// TIA Portal project "PLC_5_LINE5" (V18)

(* hardware
DEVICE "S7-1500/ET200MP station_1"  S7-1500 station
   slot 0: "Rail_0"  Rack  6ES7 590-1***0-0AA0
   slot 1: "PLC_1"  CPU 1511-1 PN  6ES7 511-1AK02-0AB0  V2.9
      slot 3: "CPU display_1"  6ES7591-1AA00-0AA0
      slot 32768: "PROFINET interface_1"  X1
         slot 32769: "Port_1"  X1 P1
         slot 32770: "Port_2"  X1 P2
      slot 34817: "Virtual CP interface port_1"  Virtual CP interface port  Virtual CP interface port
   slot 2: "DI 32x24VDC HF_1"  DI 32x24VDC HF  6ES7 521-1BL00-0AB0  V2.2
   slot 3: "DQ 32x24VDC/0.5A HF_1"  DQ 32x24VDC/0.5A HF  6ES7 522-1BL01-0AB0  V1.1
*)

// ===== PLC "PLC_1"  CPU 1511-1 PN =====

VAR_GLOBAL   // PLC tag table "Default tag table"
   "Tag_1" AT %I4.3 : Bool;
   "Tag_2" AT %I4.4 : Bool;
   "Tag_3" AT %I4.5 : Bool;
   "Tag_4" AT %I4.0 : Bool;
   "Tag_5" AT %I4.1 : Bool;
   "Tag_6" AT %I5.0 : Bool;
   "Tag_7" AT %I5.2 : Bool;
   "Tag_8" AT %I6.3 : Bool;
   "Tag_9" AT %I5.3 : Bool;
   "Tag_10" AT %I5.4 : Bool;
   "Tag_11" AT %I5.5 : Bool;
   "Tag_12" AT %I5.6 : Bool;
   "Tag_13" AT %I5.7 : Bool;
   "Tag_14" AT %I6.0 : Bool;
   "Tag_15" AT %I6.1 : Bool;
   "Tag_16" AT %I6.2 : Bool;
   "Tag_17" AT %Q1.6 : Bool;
   "Tag_18" AT %Q1.7 : Bool;
   "Tag_19" AT %Q2.0 : Bool;
   "Tag_20" AT %Q2.1 : Bool;
   "Tag_21" AT %Q2.2 : Bool;
   "Tag_22" AT %Q2.3 : Bool;
   "Tag_23" AT %I0.3 : Bool;
   "Tag_24" AT %I0.4 : Bool;
   "Tag_25" AT %I0.5 : Bool;
   "Tag_26" AT %I0.0 : Bool;
   "Tag_27" AT %I0.1 : Bool;
   "Tag_28" AT %I1.0 : Bool;
   "Tag_29" AT %I2.7 : Bool;
   "Tag_30" AT %I3.1 : Bool;
   "Tag_31" AT %I1.6 : Bool;
   "Tag_32" AT %I1.7 : Bool;
   "Tag_33" AT %I2.0 : Bool;
   "Tag_34" AT %I2.1 : Bool;
   "Tag_35" AT %I2.2 : Bool;
   "Tag_36" AT %I2.3 : Bool;
   "Tag_37" AT %I2.4 : Bool;
   "Tag_38" AT %I2.5 : Bool;
   "Tag_39" AT %I2.6 : Bool;
   "Tag_40" AT %I3.0 : Bool;
   "Tag_41" AT %Q0.4 : Bool;
   "Tag_42" AT %Q0.5 : Bool;
   "Tag_43" AT %Q0.6 : Bool;
   "Tag_44" AT %Q0.7 : Bool;
   "Tag_45" AT %Q1.0 : Bool;
   "Tag_46" AT %Q1.1 : Bool;
END_VAR

TYPE "typeTask"
   STRUCT
      station : Int;
      dwell_s : Int;
      crane : String[4];
      tank_name : String[10];
      prev : Int;
      next : Int;
      status : Int;
   END_STRUCT;
END_TYPE

TYPE "typeCraneData"
   STRUCT
      task_count : Int;
      tasks : Array[1..20] of "typeTask";
      cmd_send : Bool;
      sts_busy : Bool;
      sts_done : Bool;
      sts_step : Int;
      sts_state : Int;
      ls_at : Array[0..20] of Bool;
      ls_dip : Bool;
      ls_up : Bool;
      ls_mid : Bool;
      btn_start : Bool;
      mv_fwd : Bool;
      mv_rev : Bool;
      mv_up : Bool;
      mv_down : Bool;
      estop : Bool;
      auto : Bool;
      cmd_reset : Bool;
      cmd_stop : Bool;
      pos : Array[0..20] of Int;
   END_STRUCT;
END_TYPE

DATA_BLOCK "Crane8Data"   // DB1
{ S7_Optimized_Access := 'TRUE' }
VERSION : 0.1
BEGIN
   pos[0] := 10;
   pos[1] := 1;
   pos[2] := 2;
   pos[3] := 3;
   pos[4] := 4;
   pos[5] := 5;
   pos[6] := 6;
   pos[7] := 7;
   pos[8] := 8;
   pos[9] := 9;
END_DATA_BLOCK

DATA_BLOCK "Crane9Data"   // DB2
{ S7_Optimized_Access := 'TRUE' }
VERSION : 0.1
BEGIN
   pos[0] := 22;
   pos[1] := 21;
   pos[10] := 11;
   pos[11] := 12;
   pos[12] := 13;
   pos[13] := 14;
   pos[14] := 15;
   pos[15] := 16;
   pos[16] := 17;
   pos[17] := 18;
   pos[18] := 19;
   pos[19] := 20;
   pos[20] := 21;
END_DATA_BLOCK

DATA_BLOCK "CraneSequencer_DB"   // DB3
{ S7_Optimized_Access := 'TRUE' }
VERSION : 0.1
// stored: InstanceOfName CraneSequencer
"CraneSequencer"
BEGIN
END_DATA_BLOCK

DATA_BLOCK "CraneSequencer_DB_1"   // DB4
{ S7_Optimized_Access := 'TRUE' }
VERSION : 0.1
// stored: InstanceOfName CraneSequencer
"CraneSequencer"
BEGIN
END_DATA_BLOCK

DATA_BLOCK "Crane8_Seq_DB"   // DB5
{ S7_Optimized_Access := 'TRUE' }
VERSION : 0.1
// stored: InstanceOfName CraneSequencer
"CraneSequencer"
BEGIN
END_DATA_BLOCK

DATA_BLOCK "Crane9_Seq_DB"   // DB6
{ S7_Optimized_Access := 'TRUE' }
VERSION : 0.1
// stored: InstanceOfName CraneSequencer
"CraneSequencer"
BEGIN
END_DATA_BLOCK

FUNCTION_BLOCK "CraneSequencer"   // FB1, SCL
{ S7_Optimized_Access := 'TRUE' }
VERSION : 0.1
   VAR_IN_OUT
      d : "typeCraneData";
   END_VAR
   VAR
      state : Int;
      idx : Int;
      count : Int;
      cur : Int;
      prevSend : Bool;
      tHold : TON_TIME;
      tDwell : TON_TIME;
   END_VAR
   VAR_TEMP
      target : Int;
      arrived : Bool;
   END_VAR
BEGIN
   // ============================================================================
   //  CraneSequencer  —  GENERIC per-crane batch sequencer  (LIBRARY block)
   // ----------------------------------------------------------------------------
   //  ONE function block reused by EVERY crane on EVERY PLC. Call once per scan
   //  from OB1, passing that crane's data block as the InOut #d. No copy, no
   //  find/replace — the crane it drives is chosen entirely by which DB you pass.
   //
   //  Block type : FUNCTION BLOCK (FB), language SCL.
   //  InOut      : d : "typeCraneData"           // the whole crane interface (a DB of this UDT)
   //  Static     : state:Int, idx:Int, count:Int, cur:Int, prevSend:Bool,
   //               tHold:TON_TIME, tDwell:TON_TIME
   //  Temp       : target:Int, arrived:Bool
   //
   //  OB1 (per crane):  CraneSequencer(d := "Crane6Data")   // its own instance DB
   //                    CraneSequencer(d := "Crane7AData")
   //
   //  Stations: 0=Parking  1=Loading  2..N = tanks (tank number + 1).
   //  States : 0 IDLE · 10 GO_LOAD · 20 LOWER_LOAD · 30 WAIT_BTN · 40 LIFT_LOAD
   //           50 GO_TANK · 60 LOWER_TANK · 70 DWELL · 80 LIFT_TANK · 85 GO_PARK · 90 DONE
   //
   //  DIRECTION IS BY PHYSICAL POSITION, NOT STATION NUMBER.
   //  The plant is NOT laid out in station-number order: Parking sits WEST of Loading, and a
   //  downstream crane's Loading is a transfer tank at the far (West) end. So travel direction
   //  is decided from #d.pos[station] — the physical left→right position of each station
   //  (1 = East-most … larger = further West). TravelTo drives WEST (mv_fwd → R-West) toward a
   //  HIGHER pos, EAST (mv_rev → R-East) toward a LOWER pos. The station's arrival switch is still
   //  #d.ls_at[station]. **Set #d.pos[] per crane** — see the PLC's position-map doc.
   //
   //  COMMANDS (app/Manager writes these):
   //    cmd_send  — arm a batch (rising edge, from IDLE).
   //    cmd_stop  — EMERGENCY HOLD: kills all motion immediately, latches state 100 (STOPPED).
   //                Does NOT clear the recipe. Clear it (and Reset) to move again.
   //    cmd_reset — CLEAN/HOME: lift clear → travel to Parking → wipe the recipe → IDLE.
   //                "As if no recipe was sent, crane back at its home." PLC clears cmd_reset when done.
   //  Extra states: 100 STOPPED · 110 RESET_LIFT · 120 RESET_HOME.
   // ============================================================================

   // ---- command overrides (run BEFORE the state machine, highest priority) ----
   IF #d.cmd_stop THEN                       // immediate emergency hold (latched)
       #d.mv_fwd := FALSE;
       #d.mv_rev := FALSE;
       #d.mv_up := FALSE;
       #d.mv_down := FALSE;
       #d.sts_busy := FALSE;
       #state := 100;
   ELSIF #d.cmd_reset AND #state <> 110 AND #state <> 120 THEN   // start homing/clear (if not already)
       // Wipe the recipe IMMEDIATELY (visible at once), then home the crane.
       #d.task_count := 0;
       #d.sts_step := 0;
       #d.sts_done := FALSE;
       #d.cmd_send := FALSE;
       #idx := 0;
       #count := 0;
       #d.sts_busy := TRUE;
       #state := 110;
   END_IF;

   #d.sts_state := #state;

   CASE #state OF
       0:  // IDLE — parked, hoist up, motors off, waiting for a batch.
           #d.mv_fwd := FALSE;
           #d.mv_rev := FALSE;
           #d.mv_up := FALSE;
           #d.mv_down := FALSE;
           #d.sts_busy := FALSE;
           #d.sts_step := 0;
           IF #d.cmd_send AND NOT #prevSend AND #d.task_count > 0 THEN
               #count := #d.task_count;
               #idx := 1;
               #d.sts_done := FALSE;
               #d.sts_busy := TRUE;
               #state := 10;
           END_IF;

       10: // GO_LOAD — travel to the Loading Area (station 1).
           #d.sts_busy := TRUE;
           #target := 1;
           #arrived := "TravelTo"(target := #d.pos[#target], cur := #d.pos[#cur],
                                  atTarget := #d.ls_at[#target],
                                  fwd => #d.mv_fwd, rev => #d.mv_rev);
           IF #arrived THEN
               #cur := #target;
               #d.mv_fwd := FALSE;
               #d.mv_rev := FALSE;
               #state := 20;
           END_IF;

       20: // LOWER_LOAD — lower the hoist until the dip limit switch is made.
           #d.mv_up := FALSE;
           #d.mv_down := TRUE;
           IF #d.ls_dip THEN
               #d.mv_down := FALSE;
               #state := 30;
           END_IF;

       30: // WAIT_BTN — operator loads material, then HOLDS btn_start for 3 s.
           #tHold(IN := #d.btn_start,
                  PT := T#3S);
           IF #tHold.Q THEN
               #state := 40;
           END_IF;

       40: // LIFT_LOAD — raise the hoist clear before travelling.
           #d.mv_down := FALSE;
           #d.mv_up := TRUE;
           IF #d.ls_up THEN
               #d.mv_up := FALSE;
               #state := 50;
           END_IF;

       50: // GO_TANK — travel to THIS task's tank station (TravelTo reverses if lower).
           #d.sts_step := #idx;
           #d.tasks[#idx].status := 1;                  // running
           #target := #d.tasks[#idx].station;
           #arrived := "TravelTo"(target := #d.pos[#target], cur := #d.pos[#cur],
                                  atTarget := #d.ls_at[#target],
                                  fwd => #d.mv_fwd, rev => #d.mv_rev);
           IF #arrived THEN
               #cur := #target;
               #d.mv_fwd := FALSE;
               #d.mv_rev := FALSE;
               #state := 60;
           END_IF;

       60: // LOWER_TANK — dip into the tank until the dip limit switch is made.
           #d.mv_up := FALSE;
           #d.mv_down := TRUE;
           IF #d.ls_dip THEN
               #d.mv_down := FALSE;
               #state := 70;
           END_IF;

       70: // DWELL — hold in the tank for this task's dwell_s seconds.
           #tDwell(IN := TRUE,
                   PT := DINT_TO_TIME(INT_TO_DINT(#d.tasks[#idx].dwell_s) * 1000));
           IF #tDwell.Q THEN
               #tDwell(IN := FALSE,
                       PT := T#0S);        // reset the timer for the next tank
               #state := 80;
           END_IF;

       80: // LIFT_TANK — lift out, mark the task done, advance or finish.
           #d.mv_down := FALSE;
           #d.mv_up := TRUE;
           IF #d.ls_up THEN
               #d.mv_up := FALSE;
               #d.tasks[#idx].status := 2;              // done
               IF #idx < #count THEN
                   #idx := #idx + 1;
                   #state := 50;                        // next tank
               ELSE
                   #state := 85;                        // all tanks done
               END_IF;
           END_IF;

       85: // GO_PARK — return home to Parking (station 0).
           #target := 0;
           #arrived := "TravelTo"(target := #d.pos[#target], cur := #d.pos[#cur],
                                  atTarget := #d.ls_at[#target],
                                  fwd => #d.mv_fwd, rev => #d.mv_rev);
           IF #arrived THEN
               #cur := #target;
               #d.mv_fwd := FALSE;
               #d.mv_rev := FALSE;
               #state := 90;
           END_IF;

       90: // DONE — raise the done flag, wait for the app to acknowledge (cmd_send → FALSE).
           #d.sts_busy := FALSE;
           #d.sts_done := TRUE;
           IF NOT #d.cmd_send THEN
               #d.sts_done := FALSE;
               #d.sts_step := 0;
               #state := 0;
           END_IF;

       100: // STOPPED — emergency hold. Motors off; leaves only via Reset (cmd_reset).
           #d.mv_fwd := FALSE;
           #d.mv_rev := FALSE;
           #d.mv_up := FALSE;
           #d.mv_down := FALSE;
           #d.sts_busy := FALSE;

       110: // RESET_LIFT — raise the hoist clear before homing.
           #d.mv_down := FALSE;
           #d.mv_up := TRUE;
           IF #d.ls_up THEN
               #d.mv_up := FALSE;
               #state := 120;
           END_IF;

       120: // RESET_HOME — travel to Parking, then wipe the recipe → IDLE.
           #target := 0;
           #arrived := "TravelTo"(target := #d.pos[#target], cur := #d.pos[#cur],
                                  atTarget := #d.ls_at[#target],
                                  fwd => #d.mv_fwd, rev => #d.mv_rev);
           IF #arrived THEN
               #cur := 0;
               #d.mv_fwd := FALSE;
               #d.mv_rev := FALSE;
               #d.task_count := 0;          // "as if no recipe was sent"
               #d.sts_step := 0;
               #d.sts_done := FALSE;
               #d.sts_busy := FALSE;
               #d.cmd_send := FALSE;
               #d.cmd_reset := FALSE;      // handshake: reset complete
               #idx := 0;
               #count := 0;
               #state := 0;                 // IDLE
           END_IF;
   END_CASE;

   #prevSend := #d.cmd_send;   // edge memory (runs every scan, after the CASE)
END_FUNCTION_BLOCK

FUNCTION "IOMap" : Void   // FC1, SCL
{ S7_Optimized_Access := 'TRUE' }
VERSION : 0.1
BEGIN
   // ============================================================================
   //  IOMap  —  PLC_5 (Line 5, cranes 8 & 9)  —  real %I/%Q ↔ crane DB mirrors
   //  FUNCTION (FC), SCL, return Void, no params. Call FIRST in OB1.
   //  Addresses from docs/plc/plant-panel-layout.md (PLC_5). Station = tank.number + 1.
   //
   //  ROLES (confirmed from the plant picture, East→West):
   //    Crane 8 = ENTRY  — loads at LOAD (East end), runs 5-2…5-5, parks P-8.
   //    Crane 9 = DOWNSTREAM — picks up at TRVL-5A (West), runs DRY-5A…5-6, parks P-9.
   //  Direction is by physical position (see ./POSITION-MAP.md): mv_fwd=West, mv_rev=East.
   // ============================================================================

   // ============================ CRANE 8  (Crane8Data) — ENTRY crane ============
   //  Loads at the LOAD bay (station 1, physical East end). Tanks run West from there;
   //  Parking (P-8) sits West of its tanks.
   "Crane8Data".ls_mid := "Tag_1";      // LS_Mid_C8
   "Crane8Data".ls_up := "Tag_2";      // LS_Up_C8
   "Crane8Data".ls_dip := "Tag_3";      // LS_Down_C8
   "Crane8Data".estop := "Tag_4";      // E-Stop_SW_C8
   "Crane8Data".auto := "Tag_5";      // Auto_SW_C8
   "Crane8Data".btn_start := "Tag_6";      // UP_Pendant_C8
   "Crane8Data".ls_at[0] := "Tag_7";      // PRK-5A_C8  (Parking — station 0)
   "Crane8Data".ls_at[1] := "Tag_8";      // LOAD-5A_C8 (Loading — entry bay)  [VERIFY on Panel_5]
   "Crane8Data".ls_at[2] := "Tag_9";      // 5-2_C8    (tank 1 -> station 2)
   "Crane8Data".ls_at[3] := "Tag_10";      // INS-5A_C8 (tank 2 -> station 3)
   "Crane8Data".ls_at[4] := "Tag_11";      // 5-3_C8    (tank 3 -> station 4)
   "Crane8Data".ls_at[5] := "Tag_12";      // INS-5B_C8 (tank 4 -> station 5)
   "Crane8Data".ls_at[6] := "Tag_13";      // 5-1_C8    (tank 5 -> station 6)
   "Crane8Data".ls_at[7] := "Tag_14";      // INS-5C_C8 (tank 6 -> station 7)
   "Crane8Data".ls_at[8] := "Tag_15";      // 5-4_C8    (tank 7 -> station 8)
   "Crane8Data".ls_at[9] := "Tag_16";      // 5-5_C8    (tank 8 -> station 9)
   "Tag_17" := "Crane8Data".mv_up;          // R-Up_C8
   "Tag_18" := "Crane8Data".mv_down;        // R-Down_C8
   "Tag_19" := "Crane8Data".mv_rev;         // R-East_C8   (East = reverse / lower position)
   "Tag_20" := "Crane8Data".mv_fwd;         // R-West_C8   (West = forward / higher position)
   "Tag_21" := "Crane8Data".mv_up OR "Crane8Data".mv_down;     // R-Hoist_C8
   "Tag_22" := "Crane8Data".mv_fwd OR "Crane8Data".mv_rev;     // R-Trolley_C8

   // ============================ CRANE 9  (Crane9Data) — DOWNSTREAM =============
   //  No LOAD bay — Loading (station 1) is the transfer pickup at TRVL-5A (West end),
   //  the same switch as station 20. Its tanks run East of TRVL-5A; Parking (P-9) is
   //  the West-most box.
   "Crane9Data".ls_mid := "Tag_23";      // LS_Mid_C9
   "Crane9Data".ls_up := "Tag_24";      // LS_Up_C9
   "Crane9Data".ls_dip := "Tag_25";      // LS_Down_C9
   "Crane9Data".estop := "Tag_26";      // E-Stop_SW_C9
   "Crane9Data".auto := "Tag_27";      // Auto_SW_C9
   "Crane9Data".btn_start := "Tag_28";      // UP_Pendant_C9
   "Crane9Data".ls_at[0] := "Tag_29";      // PRK-5B_C9  (Parking — station 0)
   "Crane9Data".ls_at[1] := "Tag_30";      // TRVL-5A_C9 (Loading = transfer pickup; same as station 20)
   "Crane9Data".ls_at[10] := "Tag_31";      // DRY-5A_C9 (tank 9  -> station 10)
   "Crane9Data".ls_at[11] := "Tag_32";      // 5-12_C9   (tank 10 -> station 11)
   "Crane9Data".ls_at[12] := "Tag_33";      // INS-5E_C9 (tank 11 -> station 12)
   "Crane9Data".ls_at[13] := "Tag_34";      // 5-11_C9   (tank 12 -> station 13)
   "Crane9Data".ls_at[14] := "Tag_35";      // 5-10_C9   (tank 13 -> station 14)
   "Crane9Data".ls_at[15] := "Tag_36";      // 5-9_C9    (tank 14 -> station 15)
   "Crane9Data".ls_at[16] := "Tag_37";      // INS-5D_C9 (tank 15 -> station 16)
   "Crane9Data".ls_at[17] := "Tag_38";      // 5-8_C9    (tank 16 -> station 17)
   "Crane9Data".ls_at[18] := "Tag_39";      // 5-7_C9    (tank 17 -> station 18)
   "Crane9Data".ls_at[19] := "Tag_40";      // 5-6_C9    (tank 18 -> station 19)
   "Crane9Data".ls_at[20] := "Tag_30";      // TRVL-5A_C9 (tank 19 -> station 20; = Loading pickup)
   "Tag_41" := "Crane9Data".mv_up;          // R-Up_C9
   "Tag_42" := "Crane9Data".mv_down;        // R-Down_C9
   "Tag_43" := "Crane9Data".mv_rev;         // R-East_C9
   "Tag_44" := "Crane9Data".mv_fwd;         // R-West_C9
   "Tag_45" := "Crane9Data".mv_up OR "Crane9Data".mv_down;     // R-Hoist_C9
   "Tag_46" := "Crane9Data".mv_fwd OR "Crane9Data".mv_rev;     // R-Trolley_C9
END_FUNCTION

FUNCTION "TravelTo" : Bool   // FC2, SCL
{ S7_Optimized_Access := 'TRUE' }
VERSION : 0.1
   VAR_INPUT
      target : Int;
      cur : Int;
      atTarget : Bool;
   END_VAR
   VAR_OUTPUT
      fwd : Bool;
      rev : Bool;
   END_VAR
BEGIN
   // TravelTo — pick the travel direction toward a target station.
   // Returns TRUE when the target limit switch is already made (arrived → stop).
   #fwd := FALSE;
   #rev := FALSE;

   IF #atTarget THEN
       ;                       // arrived: leave both motors off
   ELSIF #target > #cur THEN
       #fwd := TRUE;           // higher station number → travel forward
   ELSE
       #rev := TRUE;           // lower station number → travel reverse
   END_IF;

   #TravelTo := #atTarget;
END_FUNCTION

ORGANIZATION_BLOCK "Main"   // OB1, LAD, ProgramCycle
TITLE = "Main Program Sweep (Cycle)"
{ S7_Optimized_Access := 'TRUE' }
VERSION : 0.1
   VAR_INPUT
      Initial_Call : Bool;   // Initial call of this OB
      Remanence : Bool;   // =True, if remanent data are available
   END_VAR
BEGIN

REGION Network 1
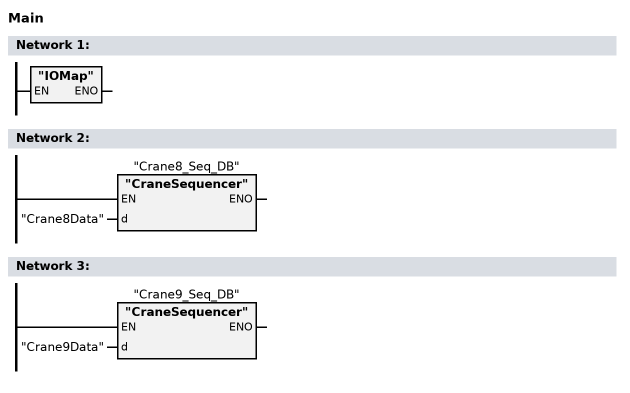
   RUNG wire#powerrail
      "IOMap"()
   END_RUNG
   // the same network as SCL:
   "IOMap"();
END_REGION

REGION Network 2
   RUNG wire#powerrail
      "Crane8_Seq_DB"(d := "Crane8Data")
   END_RUNG
   // the same network as SCL:
   "Crane8_Seq_DB"(d := "Crane8Data");   // "CraneSequencer"
END_REGION

REGION Network 3
   RUNG wire#powerrail
      "Crane9_Seq_DB"(d := "Crane9Data")
   END_RUNG
   // the same network as SCL:
   "Crane9_Seq_DB"(d := "Crane9Data");   // "CraneSequencer"
END_REGION
END_ORGANIZATION_BLOCK